// TIA Portal project "Star_Delta_Starter_V20" (V20)
// Design an automatic Star-Delta starter for a three-phase induction motor using a Siemens S7-1200 PLC. The motor shall start in Star mode, automatically transfer to Delta mode after 5 seconds, and stop immediately when the Stop button is pressed. Electrical and software interlocking shall prevent the Star and Delta contactors from being energized simultaneously.

(* hardware
DEVICE "S7-1200 station_1"  S7-1200 Station
   slot 0: "Rack_0"  S7-1200 Rack  Rack  V1.0
   slot 1: "PLC_1"  CPU 1212C DC/DC/DC  6ES7 212-1AE40-0XB0  V4.6
*)

// ===== PLC "PLC_1"  CPU 1212C DC/DC/DC =====

VAR_GLOBAL   // PLC tag table "Default tag table"
   "Start_PB" AT %I0.0 : Bool;
   "Stop_PB" AT %I0.1 : Bool;
   "Emergency_Stop" AT %I0.2 : Bool;
   "Motor_OL" AT %I0.3 : Bool;
   "Main_Contactor" AT %Q0.0 : Bool;
   "Star_Contactor" AT %Q0.1 : Bool;
   "Delta_Contactor" AT %Q0.2 : Bool;
   "Run_Lamp" AT %Q0.3 : Bool;
   "Fault_Lamp" AT %Q0.4 : Bool;
   "Motor_Run" AT %M0.0 : Bool;
   "Star_Mode" AT %M0.1 : Bool;
   "Delta_Mode" AT %M0.2 : Bool;
   "Fault" AT %M0.3 : Bool;
   "Tag_1" AT %M0.4 : Bool;
   "Tag_2" AT %M0.5 : Bool;
END_VAR

// folder: System blocks/Program resources

DATA_BLOCK "TON_Star"   // DB1
{ S7_Optimized_Access := 'TRUE' }
AUTHOR : Simatic
FAMILY : IEC
NAME : IEC_TMR
VERSION : 1.0
// stored: InstanceOfName IEC_TIMER
"IEC_TIMER"
BEGIN
END_DATA_BLOCK

DATA_BLOCK "TON_Transition"   // DB2
{ S7_Optimized_Access := 'TRUE' }
AUTHOR : Simatic
FAMILY : IEC
NAME : IEC_TMR
VERSION : 1.0
// stored: InstanceOfName IEC_TIMER
"IEC_TIMER"
BEGIN
END_DATA_BLOCK

// folder: (top level)

ORGANIZATION_BLOCK "Main"   // OB1, LAD, ProgramCycle
TITLE = "Main Program Sweep (Cycle)"
{ S7_Optimized_Access := 'TRUE' }
VERSION : 0.1
   VAR_INPUT
      Initial_Call : Bool;   // Initial call of this OB
      Remanence : Bool;   // =True, if remanent data are available
   END_VAR
BEGIN

REGION Network 1: Main_Contactor
   // S
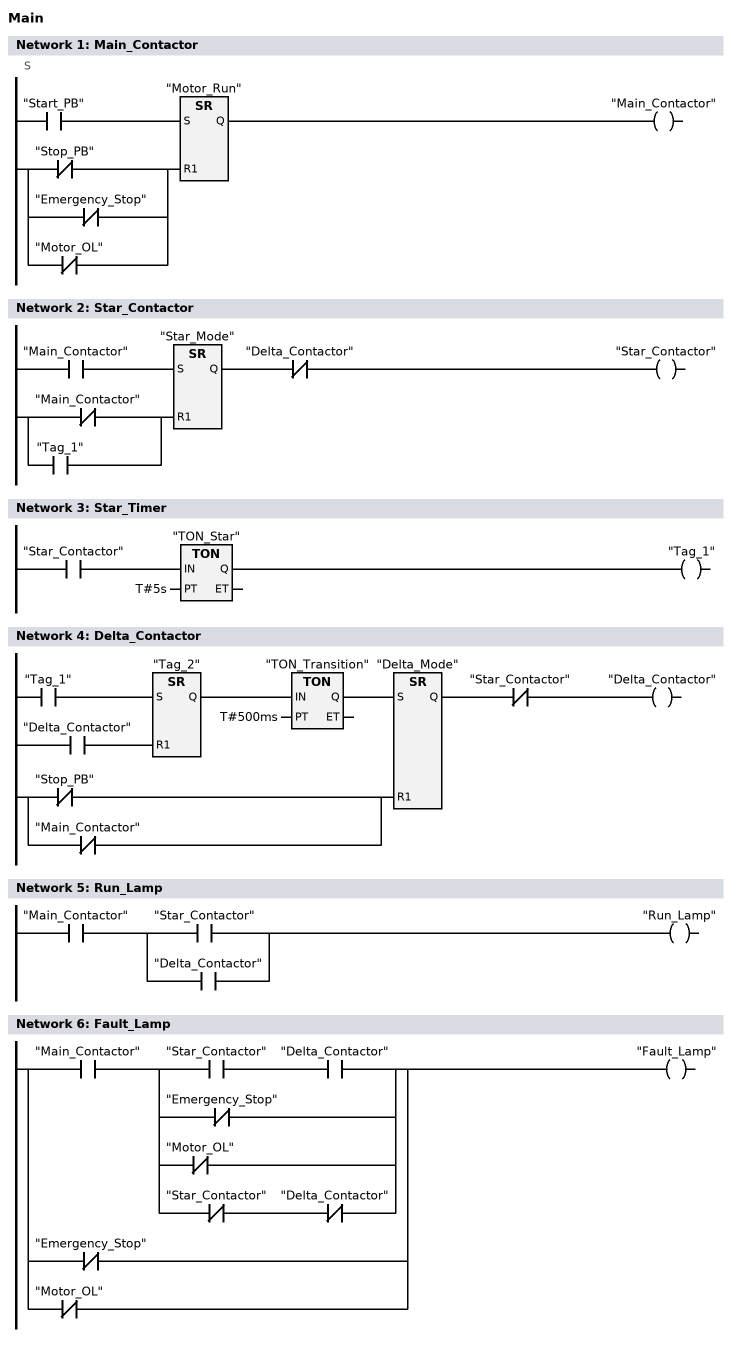
   RUNG wire#powerrail
      Contact( "Start_PB" )
      S_SR(operand := "Motor_Run", r1 := wire#w1)
      Coil( "Main_Contactor" )
   END_RUNG
   RUNG wire#powerrail
      I_Contact( "Stop_PB" )
   END_RUNG wire#w1
   RUNG wire#powerrail
      I_Contact( "Emergency_Stop" )
   END_RUNG wire#w1
   RUNG wire#powerrail
      I_Contact( "Motor_OL" )
   END_RUNG wire#w1
   // the same network as SCL:
   IF "Start_PB" THEN
       "Motor_Run" := TRUE;   // SR flip-flop
   END_IF;
   IF NOT "Stop_PB" OR NOT "Emergency_Stop" OR NOT "Motor_OL" THEN "Motor_Run" := FALSE; END_IF;
   "Main_Contactor" := "Motor_Run";
END_REGION

REGION Network 2: Star_Contactor
   RUNG wire#powerrail
      Contact( "Main_Contactor" )
      S_SR(operand := "Star_Mode", r1 := wire#w1)
      I_Contact( "Delta_Contactor" )
      Coil( "Star_Contactor" )
   END_RUNG
   RUNG wire#powerrail
      I_Contact( "Main_Contactor" )
   END_RUNG wire#w1
   RUNG wire#powerrail
      Contact( "Tag_1" )
   END_RUNG wire#w1
   // the same network as SCL:
   IF "Main_Contactor" THEN
       "Star_Mode" := TRUE;   // SR flip-flop
   END_IF;
   IF NOT "Main_Contactor" OR "Tag_1" THEN "Star_Mode" := FALSE; END_IF;
   "Star_Contactor" := "Star_Mode" AND NOT "Delta_Contactor";
END_REGION

REGION Network 3: Star_Timer
   "TON_Star".TON(IN := "Star_Contactor", PT := T#5s);
   "Tag_1" := "TON_Star".Q;
END_REGION

REGION Network 4: Delta_Contactor
   IF "Tag_1" THEN
       "Tag_2" := TRUE;   // SR flip-flop
   END_IF;
   IF "Delta_Contactor" THEN "Tag_2" := FALSE; END_IF;
   "TON_Transition".TON(IN := "Tag_2", PT := T#500ms);
   IF "TON_Transition".Q THEN
       "Delta_Mode" := TRUE;   // SR flip-flop
   END_IF;
   IF NOT "Stop_PB" OR NOT "Main_Contactor" THEN "Delta_Mode" := FALSE; END_IF;
   "Delta_Contactor" := "Delta_Mode" AND NOT "Star_Contactor";
END_REGION

REGION Network 5: Run_Lamp
   RUNG wire#powerrail
      Contact( "Main_Contactor" )
      wire#w1
      Contact( "Star_Contactor" )
      wire#w2
      Coil( "Run_Lamp" )
   END_RUNG
   RUNG wire#w1
      Contact( "Delta_Contactor" )
   END_RUNG wire#w2
   // the same network as SCL:
   "Run_Lamp" := "Main_Contactor" AND ("Star_Contactor" OR "Delta_Contactor");
END_REGION

REGION Network 6: Fault_Lamp
   RUNG wire#powerrail
      Contact( "Main_Contactor" )
      wire#w1
      Contact( "Star_Contactor" )
      Contact( "Delta_Contactor" )
      wire#w2
      Coil( "Fault_Lamp" )
   END_RUNG
   RUNG wire#w1
      I_Contact( "Emergency_Stop" )
   END_RUNG wire#w2
   RUNG wire#w1
      I_Contact( "Motor_OL" )
   END_RUNG wire#w2
   RUNG wire#w1
      I_Contact( "Star_Contactor" )
      I_Contact( "Delta_Contactor" )
   END_RUNG wire#w2
   RUNG wire#powerrail
      I_Contact( "Emergency_Stop" )
   END_RUNG wire#w2
   RUNG wire#powerrail
      I_Contact( "Motor_OL" )
   END_RUNG wire#w2
   // the same network as SCL:
   "Fault_Lamp" := ("Main_Contactor" AND (("Star_Contactor" AND "Delta_Contactor") OR NOT "Emergency_Stop" OR NOT "Motor_OL" OR (NOT "Star_Contactor" AND NOT "Delta_Contactor"))) OR NOT "Emergency_Stop" OR NOT "Motor_OL";
END_REGION
END_ORGANIZATION_BLOCK